PROGRAM Gr00MachineMode
VAR_INPUT
	(* Input variables / Eingang Variablen *)
	bEnable					:BOOL;						(* Enable Gr00MachineMode *)
END_VAR
VAR
	(* Enummerations *)

	(* Variables *)

	(* References *)

	(* Interfaces *)

	(* Instances *)

END_VAR

IF NOT bEnable
THEN
	RETURN;
END_IF;

Gr00Auto(bEnable := TRUE);			(* Call Program *)
Gr00Home(bEnable := TRUE);			(* Call Program *)
Gr00Manual(bEnable := TRUE);			(* Call Program *)

END_PROGRAM

(* stored: Version 1.1.0.1, ProductVersion 3.1.4024.15
   POU Gr00MachineMode: Id {56898725-d717-4228-bb64-052096a209f9}, SpecialFunc None *)
